SUBAPPLICATION SubApp_PC_B (* Geraet B: Methode AddValues (opcua.adoc): SERVER_1_2 + F_ADD; Input_I1 ruft sie per CLIENT_2_1 mit 43 und 10 auf (Ergebnis 53) *)
  (* Standard: 61499-2; Description: Copyright (c) 2026 Meisterschulen am Ostbahnhof This program and the accompanying materials are made available under the terms of the Eclipse Public License 2.0 which is available at https://www.eclipse.org/legal/epl-2.0/ SPDX-License-Identifier: EPL-2.0 *)
  (* Version 1.0, 2026-10-18, Franz Höpfinger, Meisterschulen am Ostbahnhof, opcua.adoc-Beispiel auf zwei Geraeten *)
  PACKAGE subapp::Training_15_OPC_UA_RES;
  IMPORT VV::const::OPC_UA::myOpcUaAddresses::T15_ADD_METHOD;
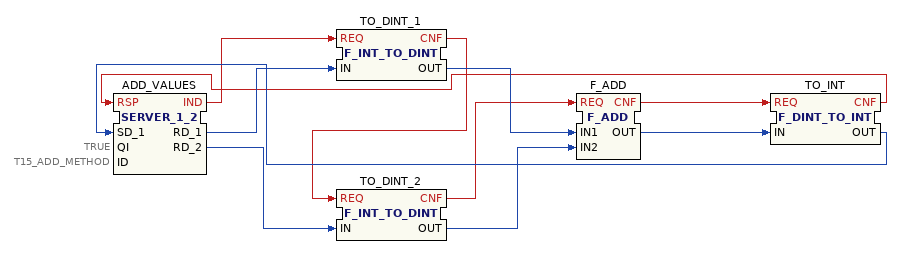
  FBS
    ADD_VALUES : iec61499::net::SERVER_1_2(QI := TRUE, ID := T15_ADD_METHOD);
    TO_DINT_1 : iec61131::conversion::F_INT_TO_DINT;
    TO_DINT_2 : iec61131::conversion::F_INT_TO_DINT;
    F_ADD : iec61131::arithmetic::F_ADD;
    TO_INT : iec61131::conversion::F_DINT_TO_INT;
  END_FBS
  EVENT_CONNECTIONS
    ADD_VALUES.IND TO TO_DINT_1.REQ;
    TO_DINT_1.CNF TO TO_DINT_2.REQ;
    TO_DINT_2.CNF TO F_ADD.REQ;
    F_ADD.CNF TO TO_INT.REQ;
    TO_INT.CNF TO ADD_VALUES.RSP;
  END_CONNECTIONS
  DATA_CONNECTIONS
    ADD_VALUES.RD_1 TO TO_DINT_1.IN;
    ADD_VALUES.RD_2 TO TO_DINT_2.IN;
    TO_DINT_1.OUT TO F_ADD.IN1;
    TO_DINT_2.OUT TO F_ADD.IN2;
    F_ADD.OUT TO TO_INT.IN;
    TO_INT.OUT TO ADD_VALUES.SD_1;
  END_CONNECTIONS
END_SUBAPPLICATION
